(* Logix 5000 project; controller lab8 vendor 1 type 14 code 149 rev 32.11; software revision 32.00 *)

TASK MainTask (continuous, watchdog 500 ms) : MainProgram

MODULES
   Local : vendor 1 type 14 code 149 (Compact 0, rev 32.11)
      Discrete_IO : Embedded (Compact 1, rev 3.1, Output RPI 20 ms)
END_MODULES

PROGRAM MainProgram   (* main routine MainRoutine *)
VAR
   LAMBER : ALIAS FOR Local:1:O.Data.1;
   LGREEN : ALIAS FOR Local:1:O.Data.2;
   LRED : ALIAS FOR Local:1:O.Data.0;
   ONS : BOOL;
   RAMBER : ALIAS FOR Local:1:O.Data.4;
   RGREEN : ALIAS FOR Local:1:O.Data.5;
   RRED : ALIAS FOR Local:1:O.Data.3;
   SENSOR : ALIAS FOR Local:1:I.Data.9;
   SENSORON : BOOL;
   start : ALIAS FOR Local:1:I.Data.2;
   START_BIT : BOOL := 1;
   STOP : ALIAS FOR Local:1:I.Data.1;
   SWITCH : BOOL := 1;
   SWITCHBIT : BOOL;
   TAMBER : TIMER := (PRE := 6000, ACC := 189, EN := 1, TT := 1);
   TGREEN : TIMER := (PRE := 9000, ACC := 9000, EN := 1, DN := 1);
   TIMER1 : TIMER := (PRE := 9000, ACC := 9000, EN := 1, DN := 1);
   TRED : TIMER := (PRE := 3000);
END_VAR

ROUTINE MainRoutine   (* ladder *)
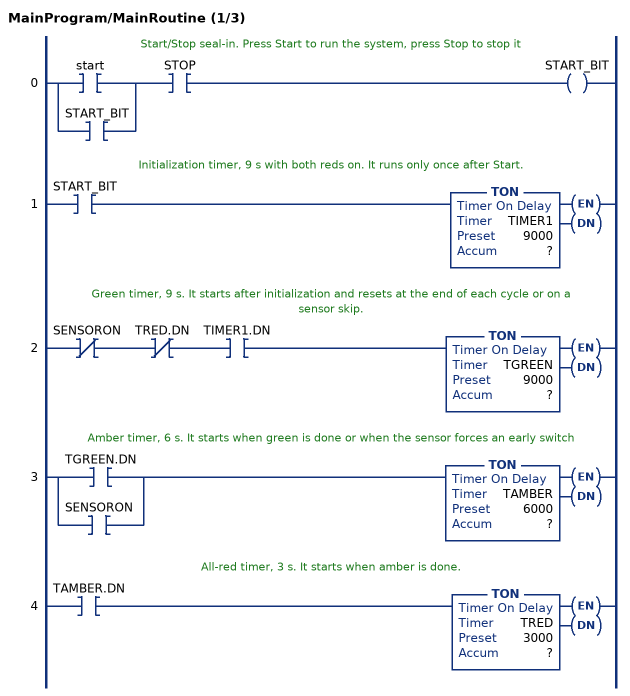
   // Start/Stop seal-in. Press Start to run the system, press Stop to stop it
   0: [XIC(start) ,XIC(START_BIT) ]XIC(STOP)OTE(START_BIT);
   // Initialization timer, 9 s with both reds on. It runs only once after Start.
   1: XIC(START_BIT)TON(TIMER1,?,?);
   // Green timer, 9 s. It starts after initialization and resets at the end of each cycle or on a sensor skip.
   2: XIO(SENSORON)XIO(TRED.DN)XIC(TIMER1.DN)TON(TGREEN,?,?);
   // Amber timer, 6 s. It starts when green is done or when the sensor forces an early switch
   3: [XIC(TGREEN.DN) ,XIC(SENSORON) ]TON(TAMBER,?,?);
   // All-red timer, 3 s. It starts when amber is done.
   4: XIC(TAMBER.DN)TON(TRED,?,?);
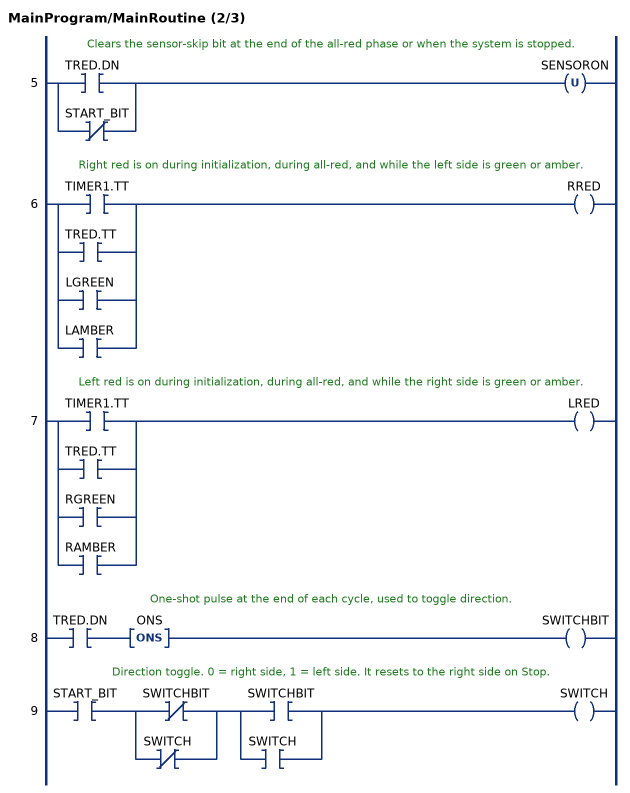
   // Clears the sensor-skip bit at the end of the all-red phase or when the system is stopped.
   5: [XIC(TRED.DN) ,XIO(START_BIT) ]OTU(SENSORON);
   // Right red is on during initialization, during all-red, and while the left side is green or amber.
   6: [[[XIC(TIMER1.TT) ,XIC(TRED.TT) ] ,XIC(LGREEN) ] ,XIC(LAMBER) ]OTE(RRED);
   // Left red is on during initialization, during all-red, and while the right side is green or amber.
   7: [[[XIC(TIMER1.TT) ,XIC(TRED.TT) ] ,XIC(RGREEN) ] ,XIC(RAMBER) ]OTE(LRED);
   // One-shot pulse at the end of each cycle, used to toggle direction.
   8: XIC(TRED.DN)ONS(ONS)OTE(SWITCHBIT);
   // Direction toggle. 0 = right side, 1 = left side. It resets to the right side on Stop.
   9: XIC(START_BIT)[XIO(SWITCHBIT) ,XIO(SWITCH) ][XIC(SWITCHBIT) ,XIC(SWITCH) ]OTE(SWITCH);
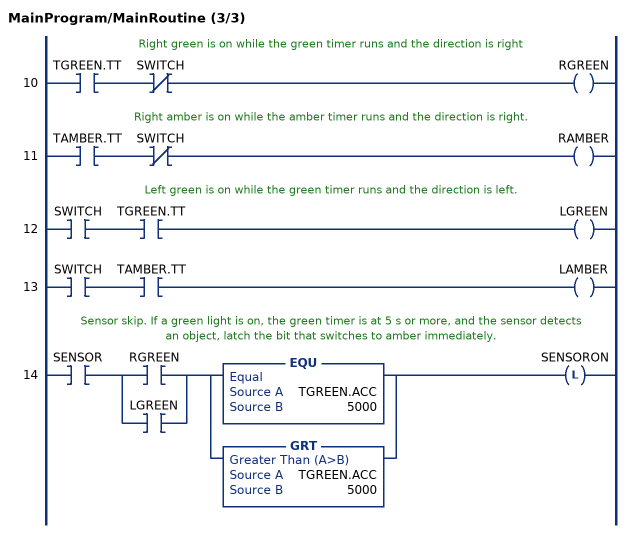
   // Right green is on while the green timer runs and the direction is right
   10: XIC(TGREEN.TT)XIO(SWITCH)OTE(RGREEN);
   // Right amber is on while the amber timer runs and the direction is right.
   11: XIC(TAMBER.TT)XIO(SWITCH)OTE(RAMBER);
   // Left green is on while the green timer runs and the direction is left.
   12: XIC(SWITCH)XIC(TGREEN.TT)OTE(LGREEN);
   13: XIC(SWITCH)XIC(TAMBER.TT)OTE(LAMBER);
   // Sensor skip. If a green light is on, the green timer is at 5 s or more, and the sensor detects an object, latch the bit that switches to amber immediately.
   14: XIC(SENSOR)[XIC(RGREEN) ,XIC(LGREEN) ][EQU(TGREEN.ACC,5000) ,GRT(TGREEN.ACC,5000) ]OTL(SENSORON);
END_ROUTINE
END_PROGRAM
